TYPE "ST_TwoHandParCfg"
VERSION : 0.1
   STRUCT
      "SchemaVersion" : UInt := 1;
      "RequireReleaseBetweenCycles" : Bool := TRUE;
   END_STRUCT;
END_TYPE
